FUNCTION_BLOCK OBSERVER_DEMO_PROCESS (* Experimental; offline checks only; native export/runtime pending *)
  (* Standard: 61499-2 *)
  (* Version 0.1, 2026-10-20, Guilherme *)
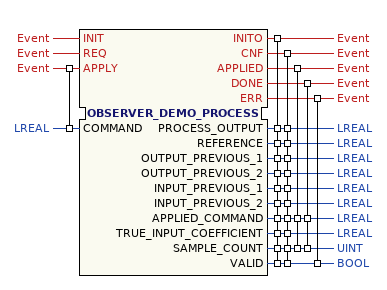
  EVENT_INPUT
    INIT;
    REQ;
    APPLY WITH COMMAND;
  END_EVENT
  EVENT_OUTPUT
    INITO WITH PROCESS_OUTPUT, REFERENCE, OUTPUT_PREVIOUS_1, OUTPUT_PREVIOUS_2, INPUT_PREVIOUS_1, INPUT_PREVIOUS_2, APPLIED_COMMAND, TRUE_INPUT_COEFFICIENT, SAMPLE_COUNT, VALID;
    CNF WITH PROCESS_OUTPUT, REFERENCE, OUTPUT_PREVIOUS_1, OUTPUT_PREVIOUS_2, INPUT_PREVIOUS_1, INPUT_PREVIOUS_2, APPLIED_COMMAND, TRUE_INPUT_COEFFICIENT, SAMPLE_COUNT, VALID;
    APPLIED WITH APPLIED_COMMAND, SAMPLE_COUNT;
    DONE WITH APPLIED_COMMAND, SAMPLE_COUNT;
    ERR WITH VALID;
  END_EVENT
  VAR_INPUT
    COMMAND : LREAL;
  END_VAR
  VAR_OUTPUT
    PROCESS_OUTPUT : LREAL;
    REFERENCE : LREAL;
    OUTPUT_PREVIOUS_1 : LREAL;
    OUTPUT_PREVIOUS_2 : LREAL;
    INPUT_PREVIOUS_1 : LREAL;
    INPUT_PREVIOUS_2 : LREAL;
    APPLIED_COMMAND : LREAL;
    TRUE_INPUT_COEFFICIENT : LREAL;
    SAMPLE_COUNT : UINT;
    VALID : BOOL;
  END_VAR
  VAR
    Y1 : LREAL;
    Y2 : LREAL;
    U1 : LREAL;
    U2 : LREAL;
    REFERENCE_COUNT : UINT;
    REFERENCE_HIGH : BOOL;
  END_VAR
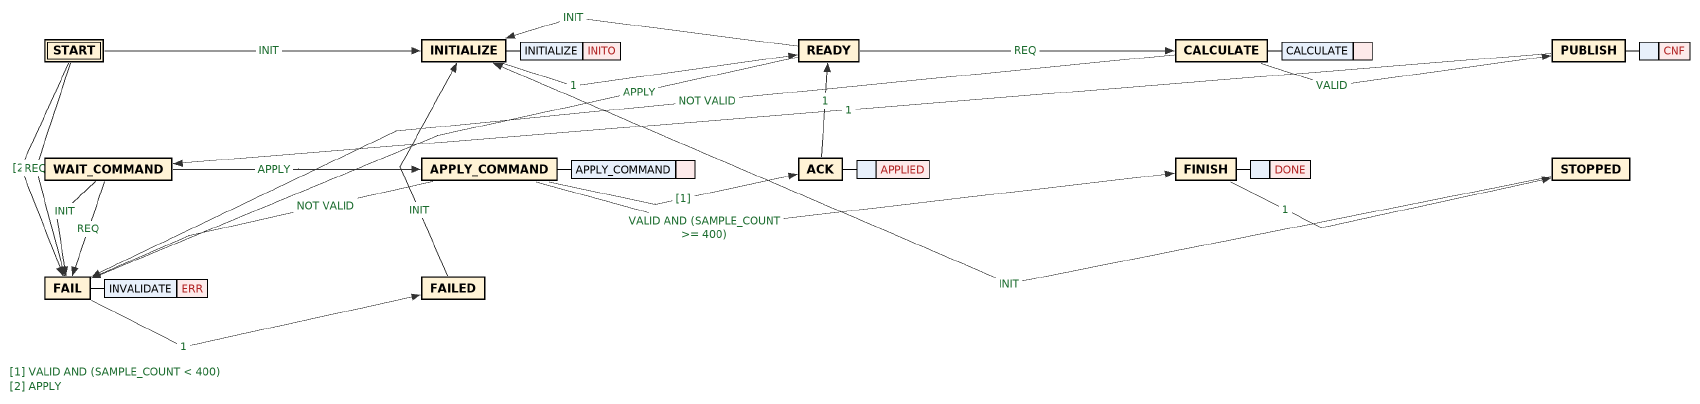
  EC_STATES
    START;
    INITIALIZE : INITIALIZE -> INITO;
    READY;
    CALCULATE : CALCULATE;
    PUBLISH : -> CNF;
    WAIT_COMMAND;
    APPLY_COMMAND : APPLY_COMMAND;
    ACK : -> APPLIED;
    FINISH : -> DONE;
    STOPPED;
    FAIL : INVALIDATE -> ERR;
    FAILED;
  END_STATES
  EC_TRANSITIONS
    START TO INITIALIZE := INIT;
    START TO FAIL := REQ;
    START TO FAIL := APPLY;
    INITIALIZE TO READY := 1;
    READY TO CALCULATE := REQ;
    READY TO INITIALIZE := INIT;
    READY TO FAIL := APPLY;
    CALCULATE TO PUBLISH := VALID;
    CALCULATE TO FAIL := NOT VALID;
    PUBLISH TO WAIT_COMMAND := 1;
    WAIT_COMMAND TO APPLY_COMMAND := APPLY;
    WAIT_COMMAND TO FAIL := REQ;
    WAIT_COMMAND TO FAIL := INIT;
    APPLY_COMMAND TO FAIL := NOT VALID;
    APPLY_COMMAND TO ACK := VALID AND (SAMPLE_COUNT < 400);
    APPLY_COMMAND TO FINISH := VALID AND (SAMPLE_COUNT >= 400);
    ACK TO READY := 1;
    FINISH TO STOPPED := 1;
    STOPPED TO INITIALIZE := INIT;
    FAIL TO FAILED := 1;
    FAILED TO INITIALIZE := INIT;
  END_TRANSITIONS
  ALGORITHM INITIALIZE IN ST:
Y1 := 0.0;
Y2 := 0.0;
U1 := 0.0;
U2 := 0.0;
PROCESS_OUTPUT := 0.0;
OUTPUT_PREVIOUS_1 := 0.0;
OUTPUT_PREVIOUS_2 := 0.0;
INPUT_PREVIOUS_1 := 0.0;
INPUT_PREVIOUS_2 := 0.0;
APPLIED_COMMAND := 0.0;
SAMPLE_COUNT := 0;
REFERENCE_COUNT := 0;
REFERENCE_HIGH := TRUE;
REFERENCE := 1.0;
TRUE_INPUT_COEFFICIENT := 0.1;
VALID := TRUE;
  END_ALGORITHM
  ALGORITHM CALCULATE IN ST:
SAMPLE_COUNT := SAMPLE_COUNT + 1;
IF REFERENCE_COUNT >= 50 THEN
REFERENCE_HIGH := NOT REFERENCE_HIGH;
REFERENCE_COUNT := 0;
END_IF;
REFERENCE_COUNT := REFERENCE_COUNT + 1;
REFERENCE := 0.8;
IF REFERENCE_HIGH THEN
REFERENCE := 1.0;
END_IF;
TRUE_INPUT_COEFFICIENT := 0.1;
IF SAMPLE_COUNT >= 151 THEN
TRUE_INPUT_COEFFICIENT := 0.4;
END_IF;
OUTPUT_PREVIOUS_1 := Y1;
OUTPUT_PREVIOUS_2 := Y2;
INPUT_PREVIOUS_1 := U1;
INPUT_PREVIOUS_2 := U2;
PROCESS_OUTPUT := 1.2 * Y1 - 0.36 * Y2 + TRUE_INPUT_COEFFICIENT * U1 + 0.06 * U2;
VALID := (PROCESS_OUTPUT >= -1.0E+100) AND (PROCESS_OUTPUT <= 1.0E+100);
  END_ALGORITHM
  ALGORITHM APPLY_COMMAND IN ST:
VALID := (COMMAND >= 0.0) AND (COMMAND <= 10.0);
IF VALID THEN
Y2 := Y1;
Y1 := PROCESS_OUTPUT;
U2 := U1;
U1 := COMMAND;
APPLIED_COMMAND := COMMAND;
END_IF;
  END_ALGORITHM
  ALGORITHM INVALIDATE IN ST:
VALID := FALSE;
  END_ALGORITHM
END_FUNCTION_BLOCK
